Omron CX-Programmer project NewProject (CX-Programmer 9.81)

# PLC NewPLC1: CJ2M CPU32
I/O table (CPU CJ2M-CPU32): rack 0 slot 11 CJ2M-EIP21

## Global symbols (name address type ; comment)
Base_at_place 2.06 BOOL  ; Base at place
Base_clamped 2.07 BOOL  ; Base clamped
Base_enable 30.03 BOOL
Base_metalic 30.01 BOOL
Base_on W30.05 BOOL  ; van valami a Base helyén
Bases_conveyor 3.06 BOOL  ; Bases conveyor
Bases_limit 2.08 BOOL  ; Pos. at limit (bases)
Clamp_base 3.07 BOOL  ; Clamp base
Clamp_lid 3.04 BOOL  ; Clamp lid
Emergency_stop 2.13 BOOL  ; Emergency stop
Grab 3.02 BOOL  ; Grab
Inductive_Base 2.14 BOOL  ; Inductive Base
Inductive_Lid 2.15 BOOL  ; Inductive Lid
Item_detected 2.02 BOOL  ; Item detected
Lid_at_place 2.03 BOOL  ; Lid at place
Lid_clamped 2.04 BOOL  ; Lid clamped
Lid_enable 30.04 BOOL
Lid_metalic 30.02 BOOL
Lids_conveyor 3.03 BOOL  ; Lids conveyor
Lids_limit 2.05 BOOL  ; Pos. at limit (lids)
Move_X 3.00 BOOL  ; Move X
Move_Z 3.01 BOOL  ; Move Z
Moving_X 2.00 BOOL  ; Moving X
Moving_Z 2.01 BOOL  ; Moving Z
Part_leaving 2.09 BOOL  ; Part leaving
Raise_bases 3.08 BOOL  ; Pos. raise (bases)
Raise_lids 3.05 BOOL  ; Pos. raise (lids)
Reset 2.11 BOOL  ; Reset
Reset_light 3.10 BOOL  ; Reset light
Start 2.10 BOOL  ; Start
Start_light 3.09 BOOL  ; Start light
Stop 2.12 BOOL  ; Stop
Stop_light 3.11 BOOL  ; Stop light
Turn 3.04 BOOL  ; Turn
base_help W4.00 BOOL
g_comp W4.03 BOOL
g_help W4.04 BOOL
g_num W5 UINT
lid_help W4.01 BOOL
m_comp W4.02 BOOL
m_help W4.05 BOOL
m_num W6 UINT
robot_enable W30.00 BOOL

## Program NewProgram1 (cyclic task 0)
Local symbols
Clamp_based BOOL
Clampe_base BOOL
Lids_enable BOOL
m_num INT
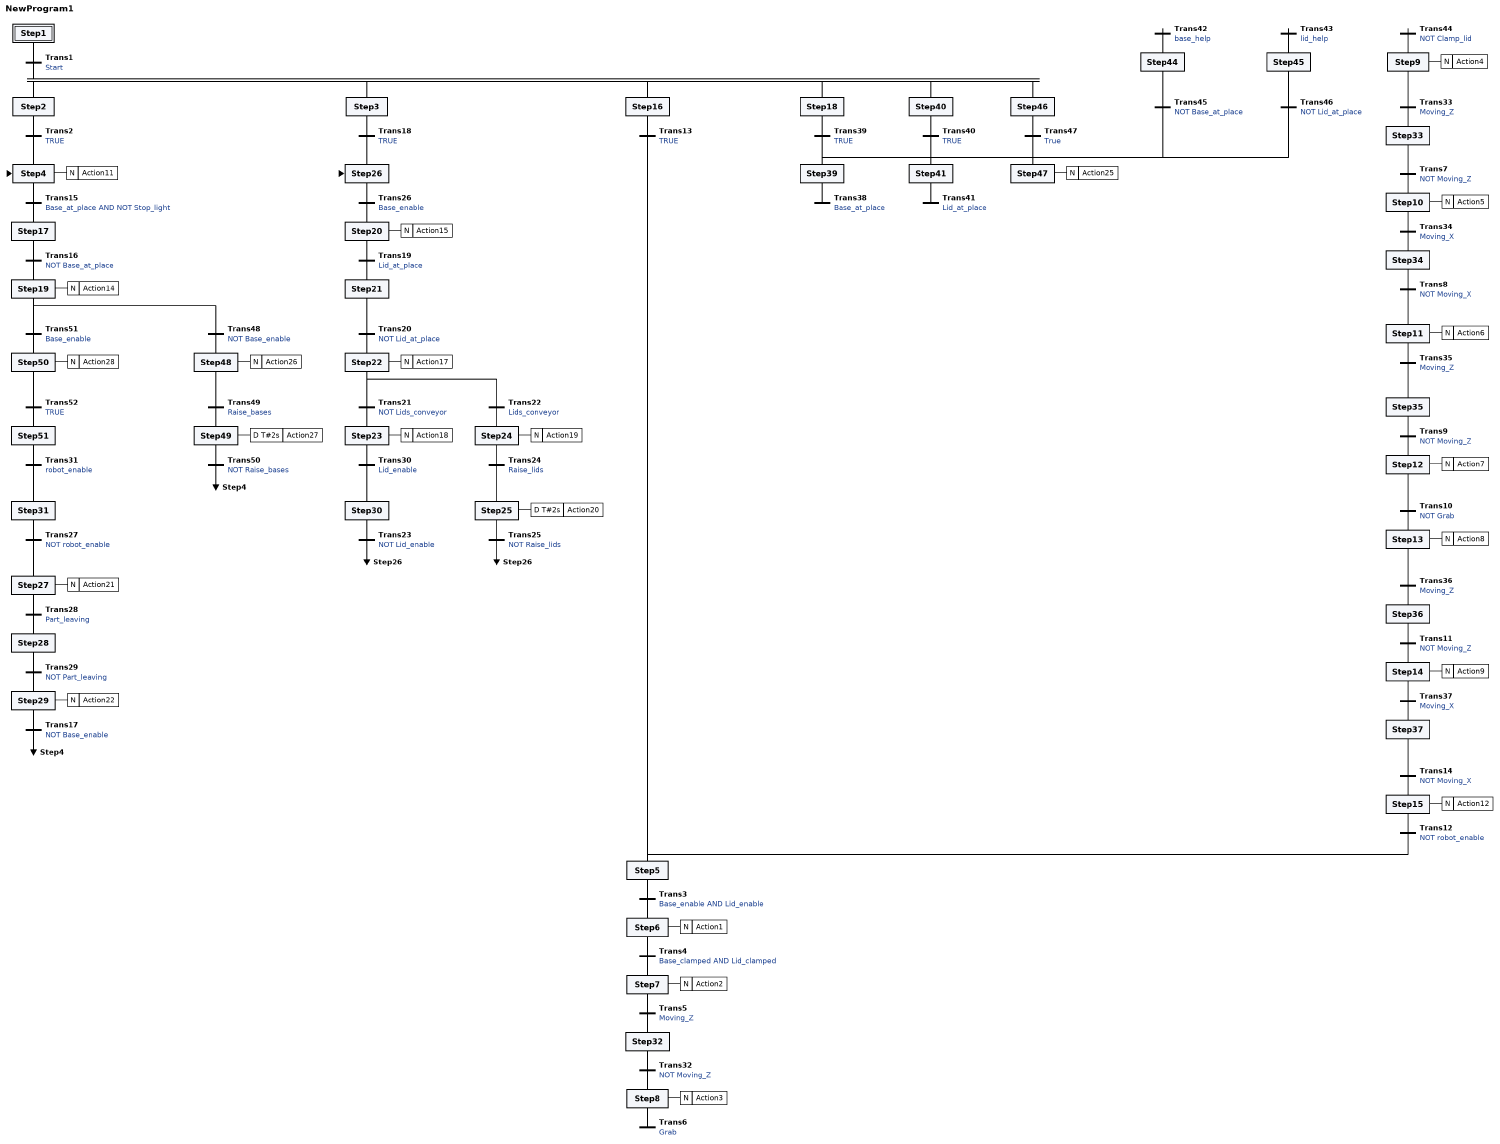
INITIAL_STEP Step1 :
END_STEP
TRANSITION Trans1 FROM Step1 TO (Step2,Step3,Step16,Step18,Step40,Step46)
 := Start;
END_TRANSITION
STEP Step2 :
END_STEP
STEP Step3 :
END_STEP
TRANSITION Trans2 FROM Step2 TO Step4
 := TRUE;
END_TRANSITION
STEP Step4 :
Action11(N) ;
END_STEP
STEP Step5 :
END_STEP
TRANSITION Trans3 FROM Step5 TO Step6
 := Base_enable AND Lid_enable;
END_TRANSITION
STEP Step6 :
Action1(N) ;
END_STEP
TRANSITION Trans4 FROM Step6 TO Step7
 := Base_clamped AND Lid_clamped;
END_TRANSITION
STEP Step7 :
Action2(N) ;
END_STEP
TRANSITION Trans5 FROM Step7 TO Step32
 := Moving_Z;
END_TRANSITION
STEP Step8 :
Action3(N) ;
END_STEP
TRANSITION Trans6 FROM Step8 TO Step43
 := Grab;
END_TRANSITION
STEP Step9 :
Action4(N) ;
END_STEP
TRANSITION Trans7 FROM Step33 TO Step10
 := NOT Moving_Z;
END_TRANSITION
STEP Step10 :
Action5(N) ;
END_STEP
TRANSITION Trans8 FROM Step34 TO Step11
 := NOT Moving_X;
END_TRANSITION
STEP Step11 :
Action6(N) ;
END_STEP
TRANSITION Trans9 FROM Step35 TO Step12
 := NOT Moving_Z;
END_TRANSITION
STEP Step12 :
Action7(N) ;
END_STEP
TRANSITION Trans10 FROM Step12 TO Step13
 := NOT Grab;
END_TRANSITION
STEP Step13 :
Action8(N) ;
END_STEP
TRANSITION Trans11 FROM Step36 TO Step14
 := NOT Moving_Z;
END_TRANSITION
STEP Step14 :
Action9(N) ;
END_STEP
TRANSITION Trans12 FROM Step15 TO Step5
 := NOT robot_enable;
END_TRANSITION
STEP Step16 :
END_STEP
TRANSITION Trans13 FROM Step16 TO Step5
 := TRUE;
END_TRANSITION
TRANSITION Trans14 FROM Step37 TO Step15
 := NOT Moving_X;
END_TRANSITION
STEP Step15 :
Action12(N) ;
END_STEP
TRANSITION Trans15 FROM Step4 TO Step17
 := Base_at_place AND NOT Stop_light;
END_TRANSITION
STEP Step17 :
END_STEP
STEP Step18 :
END_STEP
TRANSITION Trans16 FROM Step17 TO Step19
 := NOT Base_at_place;
END_TRANSITION
STEP Step19 :
Action14(N) ;
END_STEP
TRANSITION Trans17 FROM Step29 TO Step4
 := NOT Base_enable;
END_TRANSITION
TRANSITION Trans18 FROM Step3 TO Step26
 := TRUE;
END_TRANSITION
STEP Step20 :
Action15(N) ;
END_STEP
TRANSITION Trans19 FROM Step20 TO Step21
 := Lid_at_place;
END_TRANSITION
STEP Step21 :
END_STEP
TRANSITION Trans20 FROM Step21 TO Step22
 := NOT Lid_at_place;
END_TRANSITION
STEP Step22 :
Action17(N) ;
END_STEP
TRANSITION Trans21 (PRIORITY := 1) FROM Step22 TO Step23
 := NOT Lids_conveyor;
END_TRANSITION
TRANSITION Trans22 (PRIORITY := 2) FROM Step22 TO Step24
 := Lids_conveyor;
END_TRANSITION
STEP Step23 :
Action18(N) ;
END_STEP
TRANSITION Trans23 FROM Step30 TO Step26
 := NOT Lid_enable;
END_TRANSITION
STEP Step24 :
Action19(N) ;
END_STEP
TRANSITION Trans24 FROM Step24 TO Step25
 := Raise_lids;
END_TRANSITION
STEP Step25 :
Action20(D,T#2s) ;
END_STEP
TRANSITION Trans25 FROM Step25 TO Step26
 := NOT Raise_lids;
END_TRANSITION
STEP Step26 :
END_STEP
TRANSITION Trans26 FROM Step26 TO Step20
 := Base_enable;
END_TRANSITION
TRANSITION Trans27 FROM Step31 TO Step27
 := NOT robot_enable;
END_TRANSITION
STEP Step27 :
Action21(N) ;
END_STEP
TRANSITION Trans28 FROM Step27 TO Step28
 := Part_leaving;
END_TRANSITION
STEP Step28 :
END_STEP
TRANSITION Trans29 FROM Step28 TO Step29
 := NOT Part_leaving;
END_TRANSITION
STEP Step29 :
Action22(N) ;
END_STEP
TRANSITION Trans30 FROM Step23 TO Step30
 := Lid_enable;
END_TRANSITION
STEP Step30 :
END_STEP
TRANSITION Trans31 FROM Step51 TO Step31
 := robot_enable;
END_TRANSITION
STEP Step31 :
END_STEP
STEP Step32 :
END_STEP
TRANSITION Trans32 FROM Step32 TO Step8
 := NOT Moving_Z;
END_TRANSITION
TRANSITION Trans33 FROM Step9 TO Step33
 := Moving_Z;
END_TRANSITION
STEP Step33 :
END_STEP
TRANSITION Trans34 FROM Step10 TO Step34
 := Moving_X;
END_TRANSITION
STEP Step34 :
END_STEP
TRANSITION Trans35 FROM Step11 TO Step35
 := Moving_Z;
END_TRANSITION
STEP Step35 :
END_STEP
TRANSITION Trans36 FROM Step13 TO Step36
 := Moving_Z;
END_TRANSITION
STEP Step36 :
END_STEP
TRANSITION Trans37 FROM Step14 TO Step37
 := Moving_X;
END_TRANSITION
STEP Step37 :
END_STEP
TRANSITION Trans38 FROM Step39 TO Step38
 := Base_at_place;
END_TRANSITION
STEP Step38 (TIME := 100ms) :
Action16(D,T#200ms) ;
END_STEP
TRANSITION Trans39 FROM Step18 TO Step39
 := TRUE;
END_TRANSITION
STEP Step39 :
END_STEP
STEP Step40 :
END_STEP
TRANSITION Trans40 FROM Step40 TO Step41
 := TRUE;
END_TRANSITION
STEP Step41 :
END_STEP
TRANSITION Trans41 FROM Step41 TO Step42
 := Lid_at_place;
END_TRANSITION
STEP Step42 (TIME := 100ms) :
Action23(D,T#200ms) ;
END_STEP
TRANSITION Trans42 FROM Step38 TO Step44
 := base_help;
END_TRANSITION
TRANSITION Trans43 FROM Step42 TO Step45
 := lid_help;
END_TRANSITION
STEP Step43 (TIME := 100ms) :
Action24(D,T#500ms) ;
END_STEP
TRANSITION Trans44 FROM Step43 TO Step9
 := NOT Clamp_lid;
END_TRANSITION
STEP Step44 :
END_STEP
TRANSITION Trans45 FROM Step44 TO Step39
 := NOT Base_at_place;
END_TRANSITION
STEP Step45 :
END_STEP
TRANSITION Trans46 FROM Step45 TO Step41
 := NOT Lid_at_place;
END_TRANSITION
STEP Step46 :
END_STEP
TRANSITION Trans47 FROM Step46 TO Step47
 := True;
END_TRANSITION
STEP Step47 :
Action25(N) ;
END_STEP
TRANSITION Trans51 (PRIORITY := 1) FROM Step19 TO Step50
 := Base_enable;
END_TRANSITION
TRANSITION Trans48 (PRIORITY := 2) FROM Step19 TO Step48
 := NOT Base_enable;
END_TRANSITION
STEP Step48 :
Action26(N) ;
END_STEP
TRANSITION Trans49 FROM Step48 TO Step49
 := Raise_bases;
END_TRANSITION
STEP Step49 :
Action27(D,T#2s) ;
END_STEP
TRANSITION Trans50 FROM Step49 TO Step4
 := NOT Raise_bases;
END_TRANSITION
STEP Step50 :
Action28(N) ;
END_STEP
TRANSITION Trans52 FROM Step50 TO Step51
 := TRUE;
END_TRANSITION
STEP Step51 :
END_STEP

### Action Action1

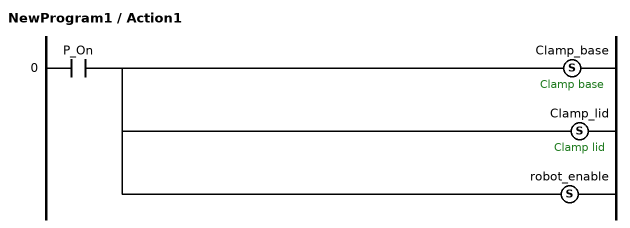
; rung 0
LD P_On
SET Clamp_base  ; Clamp base
SET Clamp_lid  ; Clamp lid
SET robot_enable

### Action Action2

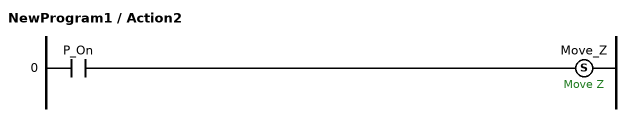
; rung 0
LD P_On
SET Move_Z  ; Move Z

### Action Action3

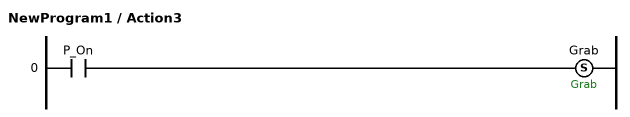
; rung 0
LD P_On
SET Grab  ; Grab

### Action Action4

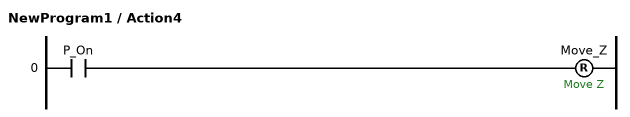
; rung 0
LD P_On
RSET Move_Z  ; Move Z

### Action Action5

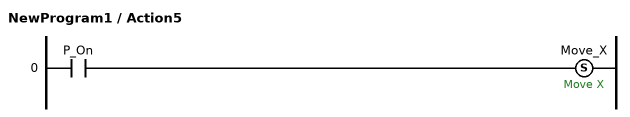
; rung 0
LD P_On
SET Move_X  ; Move X

### Action Action6

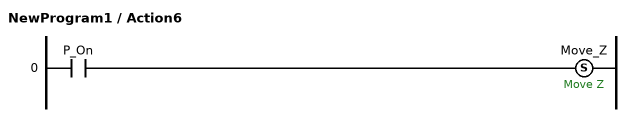
; rung 0
LD P_On
SET Move_Z  ; Move Z

### Action Action7

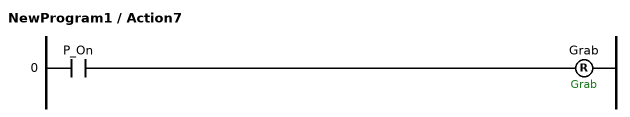
; rung 0
LD P_On
RSET Grab  ; Grab

### Action Action8

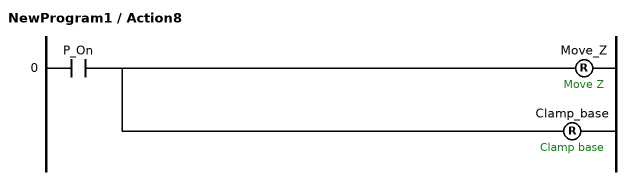
; rung 0
LD P_On
RSET Move_Z  ; Move Z
RSET Clamp_base  ; Clamp base

### Action Action9

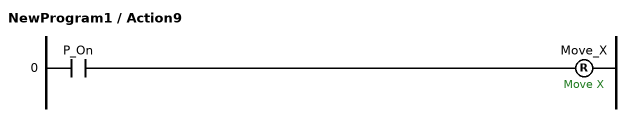
; rung 0
LD P_On
RSET Move_X  ; Move X

### Action Action10

### Action Action12

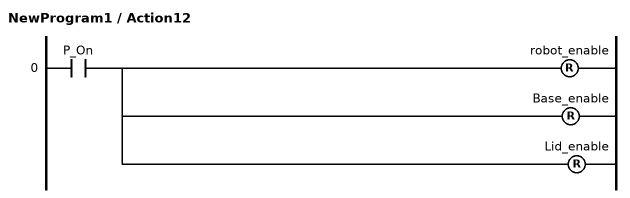
; rung 0
LD P_On
RSET robot_enable
RSET Base_enable
RSET Lid_enable

### Action Action11

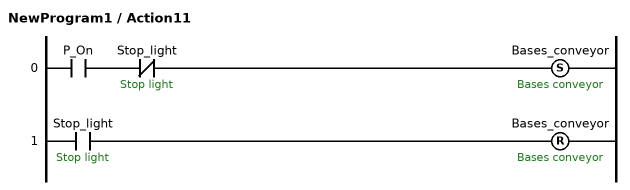
; rung 0
LD P_On
ANDNOT Stop_light  ; Stop light
SET Bases_conveyor  ; Bases conveyor
; rung 1
LD Stop_light  ; Stop light
RSET Bases_conveyor  ; Bases conveyor

### Action Action13

### Action Action14

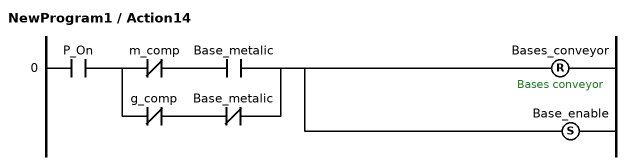
; rung 0
LD P_On
LDNOT m_comp
AND Base_metalic
LDNOT g_comp
ANDNOT Base_metalic
ORLD
ANDLD
RSET Bases_conveyor  ; Bases conveyor
SET Base_enable

### Action Action15

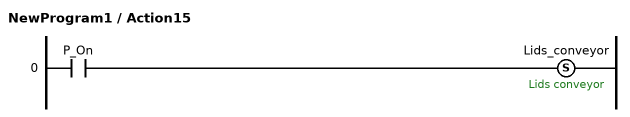
; rung 0
LD P_On
SET Lids_conveyor  ; Lids conveyor

### Action Action17

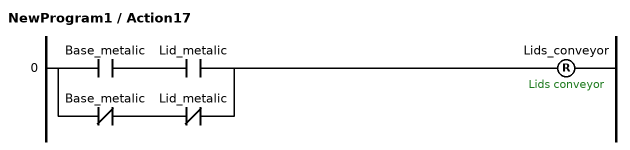
; rung 0
LD Base_metalic
AND Lid_metalic
LDNOT Base_metalic
ANDNOT Lid_metalic
ORLD
RSET Lids_conveyor  ; Lids conveyor

### Action Action18

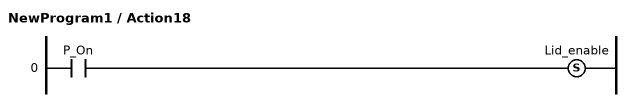
; rung 0
LD P_On
SET Lid_enable

### Action Action19

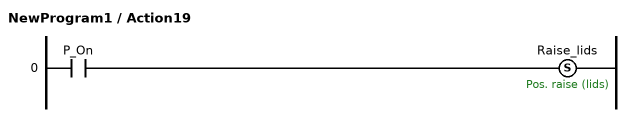
; rung 0
LD P_On
SET Raise_lids  ; Pos. raise (lids)

### Action Action20

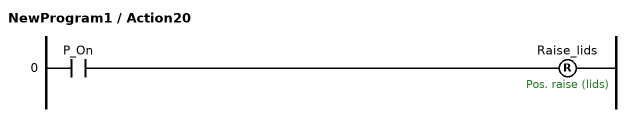
; rung 0
LD P_On
RSET Raise_lids  ; Pos. raise (lids)

### Action Action21

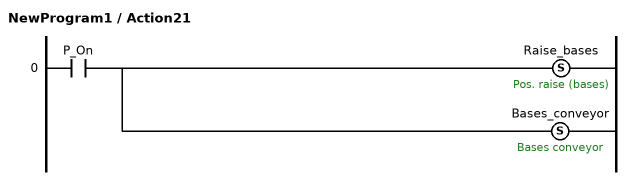
; rung 0
LD P_On
SET Raise_bases  ; Pos. raise (bases)
SET Bases_conveyor  ; Bases conveyor

### Action Action22

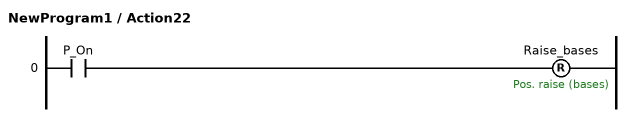
; rung 0
LD P_On
RSET Raise_bases  ; Pos. raise (bases)

### Action Action16

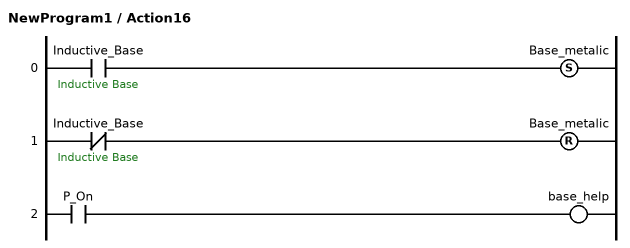
; rung 0
LD Inductive_Base  ; Inductive Base
SET Base_metalic
; rung 1
LDNOT Inductive_Base  ; Inductive Base
RSET Base_metalic
; rung 2
LD P_On
OUT base_help

### Action Action23

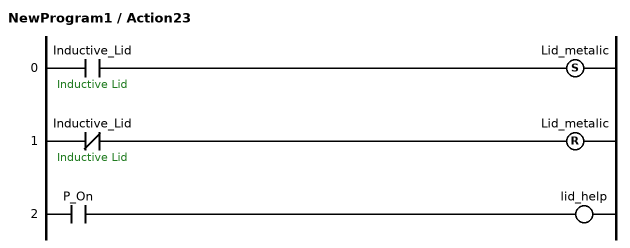
; rung 0
LD Inductive_Lid  ; Inductive Lid
SET Lid_metalic
; rung 1
LDNOT Inductive_Lid  ; Inductive Lid
RSET Lid_metalic
; rung 2
LD P_On
OUT lid_help

### Action Action24

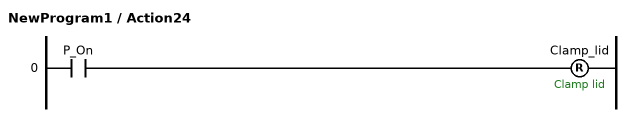
; rung 0
LD P_On
RSET Clamp_lid  ; Clamp lid

### Action Action25

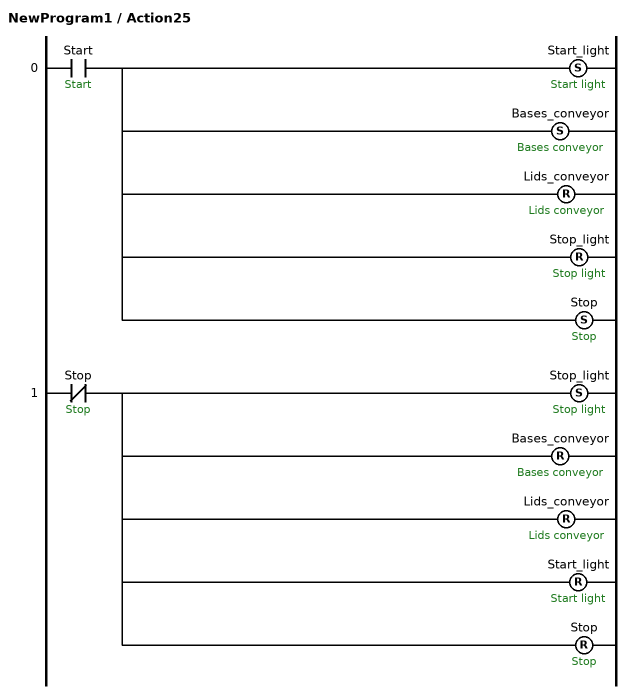
; rung 0
LD Start  ; Start
SET Start_light  ; Start light
SET Bases_conveyor  ; Bases conveyor
RSET Lids_conveyor  ; Lids conveyor
RSET Stop_light  ; Stop light
SET Stop  ; Stop
; rung 1
LDNOT Stop  ; Stop
SET Stop_light  ; Stop light
RSET Bases_conveyor  ; Bases conveyor
RSET Lids_conveyor  ; Lids conveyor
RSET Start_light  ; Start light
RSET Stop  ; Stop

### Action Action26

